// TIA Portal V21 export
// export: Created 2026-11-09T01:07:07.9028886Z, ExportSetting WithDefaults, DisplayName Totally Integrated Automation Portal, DisplayVersion V21 Update 3, DisplayName STEP 7 Professional, DisplayVersion V21 Update 3, DisplayName STEP 7 Safety, DisplayVersion V21, DisplayName Tech WebApplication, DisplayVersion V21, DisplayName WinCC Basic/Comfort/Advanced, DisplayVersion V21 Update 3, DisplayName WinCC Unified, DisplayVersion V21 Update 3
FUNCTION "FC_Typed" : Int   // FC1, SCL
{ S7_Optimized_Access := 'TRUE' }
// stored: AutoNumber true, IsIECCheckEnabled false, SetENOAutomatically false, UDAEnableTagReadback false
   VAR_INPUT
      "a" : Int;
      "b" : Int;
   END_VAR
BEGIN
   #FC_Typed := #a * #b;
END_FUNCTION
